TYPE ST_Mess_Logger :
STRUCT
	iErNum					: INT;
	sTime					: STRING[20];
	sDate					: STRING[20];
	sDescription				: STRING[40];
END_STRUCT
END_TYPE

(* stored: Version 1.1.0.1, ProductVersion 3.1.4024.13
   DUT ST_Mess_Logger: Id {7ecf682e-548d-47f1-ad95-4b836eb6574e} *)
